// TIA Portal V21 export
Screen "T05_BtnInv"  1024x768, Number=25
  ScreenLayer 
    Button "P_BtnInv" at 0,0 size 100x30  TextOff="BTN", TextOn="BTN"
      EventHandler   EventType=Press
        FunctionCall "InvertBit"
          FunctionParameter "Tag"  Tag=SwOn
